{attribute 'qualified_only'}
TYPE XtsMoverDetectionState :
(
	WaitingForCommandStart := 0,
	SetATrackForDetection := 1,                                              
	TriggeringRedetection := 2,
	WaitingForAllMoversValid := 3,                                 
	CheckingAllMoverFound := 4,
	TriggeringMoverIdDetection := 9,
	MoverDetectionFault := 99
);
END_TYPE

(* stored: Version 1.1.0.1
   DUT XtsMoverDetectionState: Id {3651fba9-c72e-488e-9f30-9cd847bba8bf} *)
